Fanuc KAREL source: KT00491.KL

PROGRAM KT00491
%NOLOCKGROUP
VAR
  P1: POSITION
  P2: JOINTPOS
  OUT: XYZWPREXT
BEGIN
  OUT = P1 : P2
END KT00491
